Universal Robots PolyScope program: pick_and_place.urp

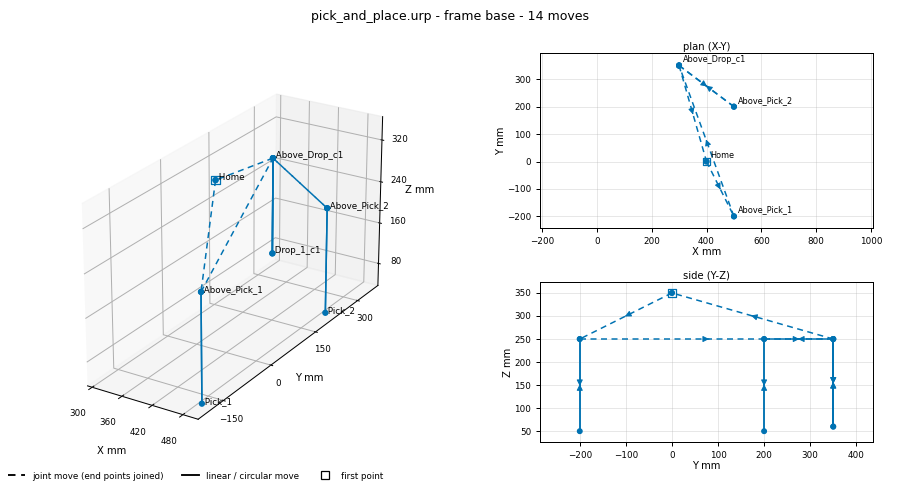
[picture p0: tool path of pick_and_place.urp in frame base, 14 of 14 moves have a stored position in this frame; points joined in program order, loops and branches not executed]
Program pick_and_place (installation=default directory=/ursim/programs createdIn=3.15.8.106339 lastSavedIn=3.15.8.106339 robotSerialNumber=2018359999)
Calibrated DH parameters: a=[0, -0.425, -0.39225, 0, 0, 0]; d=[0.089159, 0, 0, 0.10915, 0.09465, 0.0823]; alpha=[1.570796, 0, 0, 1.570796, -1.570796, 0]; deltaTheta=[0, 0, 0, 0, 0, 0]
Robot Program (runOnlyOnce=true)
  Set DigitalOutput (payload=0 tcpAsCog=true) pin=digital_out[0]; digitalValue=0
  MoveJ speed 60 deg/s, acceleration 80 deg/s^2 (useActiveTCP=true)
    Waypoint Home: TCP in base x=400 y=0 z=350 mm, rx=0 ry=3.1416 rz=0 rad; joints [15.835, -77, -113.424, -79.577, 90, 105.835] deg
  Loop Forever
    MoveJ speed 60 deg/s, acceleration 80 deg/s^2 (useActiveTCP=true)
      Waypoint Above_Pick_1: TCP in base x=500 y=-200 z=250 mm, rx=0 ry=3.1416 rz=0 rad; joints [-10.107, -101.009, -105.33, -63.661, 90, 79.893] deg
    Wait Sleep waitTime=0.3
    MoveL speed 250 mm/s, acceleration 500 mm/s^2 (useActiveTCP=true) feature=Base
      Waypoint Pick_1: TCP in base x=500 y=-200 z=50 mm, rx=0 ry=3.1416 rz=0 rad; joints [-10.107, -120.037, -115.856, -34.107, 90, 79.893] deg
    Set DigitalOutput (payload=1 tcpAsCog=true) pin=digital_out[0]; digitalValue=1
    Wait Sleep waitTime=0.5
    MoveL speed 250 mm/s, acceleration 500 mm/s^2 (useActiveTCP=true) feature=Base
      Waypoint Above_Pick_1_ret: TCP in base x=500 y=-200 z=250 mm, rx=0 ry=3.1416 rz=0 rad; joints [-10.107, -101.009, -105.33, -63.661, 90, 79.893] deg
    MoveJ speed 60 deg/s, acceleration 80 deg/s^2 (useActiveTCP=true)
      Waypoint Above_Drop_c1: TCP in base x=300 y=350 z=250 mm, rx=0 ry=3.1416 rz=0 rad; joints [63.095, -90.762, -116.853, -62.385, 90, 153.095] deg
    Wait Sleep waitTime=0.3
    MoveL speed 250 mm/s, acceleration 500 mm/s^2 (useActiveTCP=true) feature=Base
      Waypoint Drop_1_c1: TCP in base x=300 y=350 z=60 mm, rx=0 ry=3.1416 rz=0 rad; joints [63.095, -112, -128.356, -29.644, 90, 153.095] deg
    Set DigitalOutput (payload=0 tcpAsCog=true) pin=digital_out[0]; digitalValue=0
    Wait Sleep waitTime=0.5
    MoveL speed 250 mm/s, acceleration 500 mm/s^2 (useActiveTCP=true) feature=Base
      Waypoint Above_Drop_c1_ret: TCP in base x=300 y=350 z=250 mm, rx=0 ry=3.1416 rz=0 rad; joints [63.095, -90.762, -116.853, -62.385, 90, 153.095] deg
    MoveJ speed 60 deg/s, acceleration 80 deg/s^2 (useActiveTCP=true)
      Waypoint Above_Pick_2: TCP in base x=500 y=200 z=250 mm, rx=0 ry=3.1416 rz=0 rad; joints [33.495, -101.009, -105.33, -63.661, 90, 123.495] deg
    Wait Sleep waitTime=0.3
    MoveL speed 250 mm/s, acceleration 500 mm/s^2 (useActiveTCP=true) feature=Base
      Waypoint Pick_2: TCP in base x=500 y=200 z=50 mm, rx=0 ry=3.1416 rz=0 rad; joints [33.495, -120.037, -115.856, -34.107, 90, 123.495] deg
    Set DigitalOutput (payload=1 tcpAsCog=true) pin=digital_out[0]; digitalValue=1
    Wait Sleep waitTime=0.5
    MoveL speed 250 mm/s, acceleration 500 mm/s^2 (useActiveTCP=true) feature=Base
      Waypoint Above_Pick_2_ret: TCP in base x=500 y=200 z=250 mm, rx=0 ry=3.1416 rz=0 rad; joints [33.495, -101.009, -105.33, -63.661, 90, 123.495] deg
    MoveJ speed 60 deg/s, acceleration 80 deg/s^2 (useActiveTCP=true)
      Waypoint Above_Drop_c2: TCP in base x=300 y=350 z=250 mm, rx=0 ry=3.1416 rz=0 rad; joints [63.095, -90.762, -116.853, -62.385, 90, 153.095] deg
    Wait Sleep waitTime=0.3
    MoveL speed 250 mm/s, acceleration 500 mm/s^2 (useActiveTCP=true) feature=Base
      Waypoint Drop_1_c2: TCP in base x=300 y=350 z=60 mm, rx=0 ry=3.1416 rz=0 rad; joints [63.095, -112, -128.356, -29.644, 90, 153.095] deg
    Set DigitalOutput (payload=0 tcpAsCog=true) pin=digital_out[0]; digitalValue=0
    Wait Sleep waitTime=0.5
    MoveL speed 250 mm/s, acceleration 500 mm/s^2 (useActiveTCP=true) feature=Base
      Waypoint Above_Drop_c2_ret: TCP in base x=300 y=350 z=250 mm, rx=0 ry=3.1416 rz=0 rad; joints [63.095, -90.762, -116.853, -62.385, 90, 153.095] deg
    MoveJ speed 60 deg/s, acceleration 80 deg/s^2 (useActiveTCP=true)
      Waypoint Home_fin: TCP in base x=400 y=0 z=350 mm, rx=0 ry=3.1416 rz=0 rad; joints [15.835, -77, -113.424, -79.577, 90, 105.835] deg
    Wait DigitalInput pin=digital_in[0]; digitalValue=1
